(* IEC 61131-3 sources: kns-port-domestic/upstream/plc-process-lib/src/Interfaces/I_AlarmSource, 1 file *)

(* ---- GetAlarm.method.decl.st ---- *)
// Тревога слота uiIndex; вне 0..AlarmCount-1 — 0
METHOD GetAlarm : I_Alarm
VAR_INPUT
    uiIndex : UINT;   // номер слота
END_VAR
